Yaskawa INFORM job: TEAM2V2.JBI

/JOB
//NAME TEAM2V2
//POS
///NPOS 25,0,25,0,0,0
///TOOL 0
///POSTYPE PULSE
///PULSE
C00000=-947,-55524,-59539,-219,-89999,0
C00001=-14550,35752,-9918,-1666,-46835,4504
C00002=-14550,47390,-9918,-1666,-46835,4504
C00003=-14208,46659,-14977,-1765,-43895,4451
C00004=-19701,43642,-20432,-2235,-40990,-11434
C00005=-19701,43642,-20432,-2235,-40990,-11434
C00006=-13594,46848,-14975,-1487,-43513,728
C00007=325,30497,-44182,13981,-25939,22710
C00008=21917,8400,-41377,7972,-38642,30634
C00009=1813,-26553,-79211,-1109,-5827,4862
C00010=1813,-26553,-79210,-1109,-5825,4862
C00011=-13828,10438,-65699,5058,-1053,2039
C00012=-14008,16266,-68247,1762,5093,3588
C00013=-13949,16746,-68323,1395,5510,3745
C00014=-20003,17976,-66586,25043,5725,-5712
C00015=-20831,-9039,-52276,8990,-15029,-1550
C00016=-20831,-9039,-52276,8990,-15029,-1550
C00017=-24056,-21474,-63521,2858,-16442,1957
C00018=-54933,3456,-76445,73932,61358,-37474
C00019=-52302,46474,-77834,59857,73358,-21814
C00020=-52409,46839,-77304,59949,73309,-21853
C00021=-55538,45410,-82065,61547,74272,-20901
C00022=-57801,33009,-87685,64436,71959,-23280
C00023=-25442,-290,-95405,25953,33870,-5925
C00024=-946,-55528,-59541,-218,-89999,0
EC00000=-1645
EC00001=-1645
EC00002=-1645
EC00003=-1645
EC00004=-1645
EC00005=-1645
EC00006=-1645
EC00007=-1645
EC00008=-1645
EC00009=-1645
EC00010=-1645
EC00011=-83284
EC00012=-83284
EC00013=-83284
EC00014=-83284
EC00015=-83284
EC00016=-164958
EC00017=-164958
EC00018=-162295
EC00019=-162295
EC00020=-162297
EC00021=-162297
EC00022=-162295
EC00023=-162295
EC00024=-1645
//INST
///DATE 2025/11/03 18:03
///ATTR SC,RW
///GROUP1 RB1,ST1
NOP
MOVJ C00000 EC00000 VJ=25.00
MOVJ C00001 EC00001 VJ=5.00
MOVJ C00002 EC00002 VJ=1.00
MOVL C00003 EC00003 V=8.3
MOVL C00004 EC00004 V=11.7
ARCON ASF#(1)
MOVC C00005 EC00005 V=50.0
MOVC C00006 EC00006 V=11.0
MOVC C00007 EC00007 V=50.0
ARCOF AEF#(1)
MOVJ C00008 EC00008 VJ=25.00
MOVJ C00009 EC00009 VJ=25.00
MOVJ C00010 EC00010 VJ=25.00
MOVJ C00011 EC00011 VJ=25.00
MOVL C00012 EC00012 V=11.0
ARCON ASF#(1)
MOVL C00013 EC00013 V=11.0
MOVL C00014 EC00014 V=11.0
ARCOF AEF#(1)
MOVJ C00015 EC00015 VJ=5.00
MOVJ C00016 EC00016 VJ=10.00
MOVJ C00017 EC00017 VJ=5.00
MOVJ C00018 EC00018 VJ=5.00
MOVL C00019 EC00019 V=50.0
MOVL C00020 EC00020 V=50.0
ARCON ASF#(1)
MOVL C00021 EC00021 V=50.0
ARCOF AEF#(1)
MOVJ C00022 EC00022 VJ=5.00
MOVJ C00023 EC00023 VJ=25.00
MOVJ C00024 EC00024 VJ=25.00
END
